ABB RAPID module: Felisac.mod

MODULE Felisac
	TASK PERS tooldata Hfeli:=[TRUE,[[85.795,-0.16,81.2],[0.819152044,0,0.573576436,0]],[1,[0,0,1],[1,0,0,0],0,0,0]];
	TASK PERS wobjdata Wfeli:=[FALSE,TRUE,"",[[0,0,0],[1,0,0,0]],[[592.85,-241.657,124.334],[0.00174513,0.00767284,-0.999953,-0.00564666]]];

ENDMODULE
